FUNCTION_BLOCK EQ_Template (* TEMPLATE for your equipment block, EQ_<Equipment>: copy it under that name, then change what says YOUR OWN, and this comment; keep the rest as it is. An equipment block: the only block that touches this equipment's pins. Skills send it what to switch over a local channel; it switches the outputs (off first, then on), reads the inputs every cycle and reports them to the skills and to OPC UA. One skill holds it at a time; on release or when the module aborts it switches everything off. Technical: A piece of equipment to make your own: one input, one output, one command besides Stop; equipment IO: owns its IO points, writes the output values its holder sends, reads its inputs every cycle and reports changes *)
  (* Standard: 61499-2 *)
  (* Version 0.1, 2026-09-28, Project contributors, AAU Smart Production Lab *)
  PACKAGE stoppering;
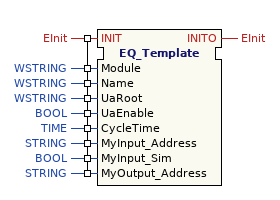
  EVENT_INPUT
    INIT : EInit WITH Module, Name, UaRoot, UaEnable, CycleTime, MyInput_Address, MyInput_Sim, MyOutput_Address; (* Initialise, once at start-up (the INIT chain); takes the values given with it *)
  END_EVENT
  EVENT_OUTPUT
    INITO : EInit; (* Initialised: the next block of the INIT chain goes on *)
  END_EVENT
  VAR_INPUT
    Module : WSTRING; (* The module's name; its local channels are named after it (loc[<Module>/...]) *)
    Name : WSTRING := "Template"; (* YOUR OWN, your equipment's name. The equipment item's name: its local channels and OPC UA folder *)
    UaRoot : WSTRING; (* The module's OPC UA folder, e.g. /Objects/Filling *)
    UaEnable : BOOL; (* Publish on OPC UA *)
    CycleTime : TIME := T#50ms; (* How often the inputs are read *)
    MyInput_Address : STRING; (* YOUR OWN, one per input pin. Where MyInput is: 'gpio[chip:line(:pull_up|:pull_down)(:active_low)]', 'pwm[chip:channel:period_ns]', 'modbus[...]', 'sim', or an IO handle's name; empty: not connected *)
    MyInput_Sim : BOOL := FALSE; (* YOUR OWN, one per input pin. The value of MyInput when simulated (address 'sim') *)
    MyOutput_Address : STRING; (* YOUR OWN, one per output pin. Where MyOutput is: 'gpio[chip:line(:pull_up|:pull_down)(:active_low)]', 'pwm[chip:channel:period_ns]', 'modbus[...]', 'sim', or an IO handle's name; empty: not connected *)
  END_VAR
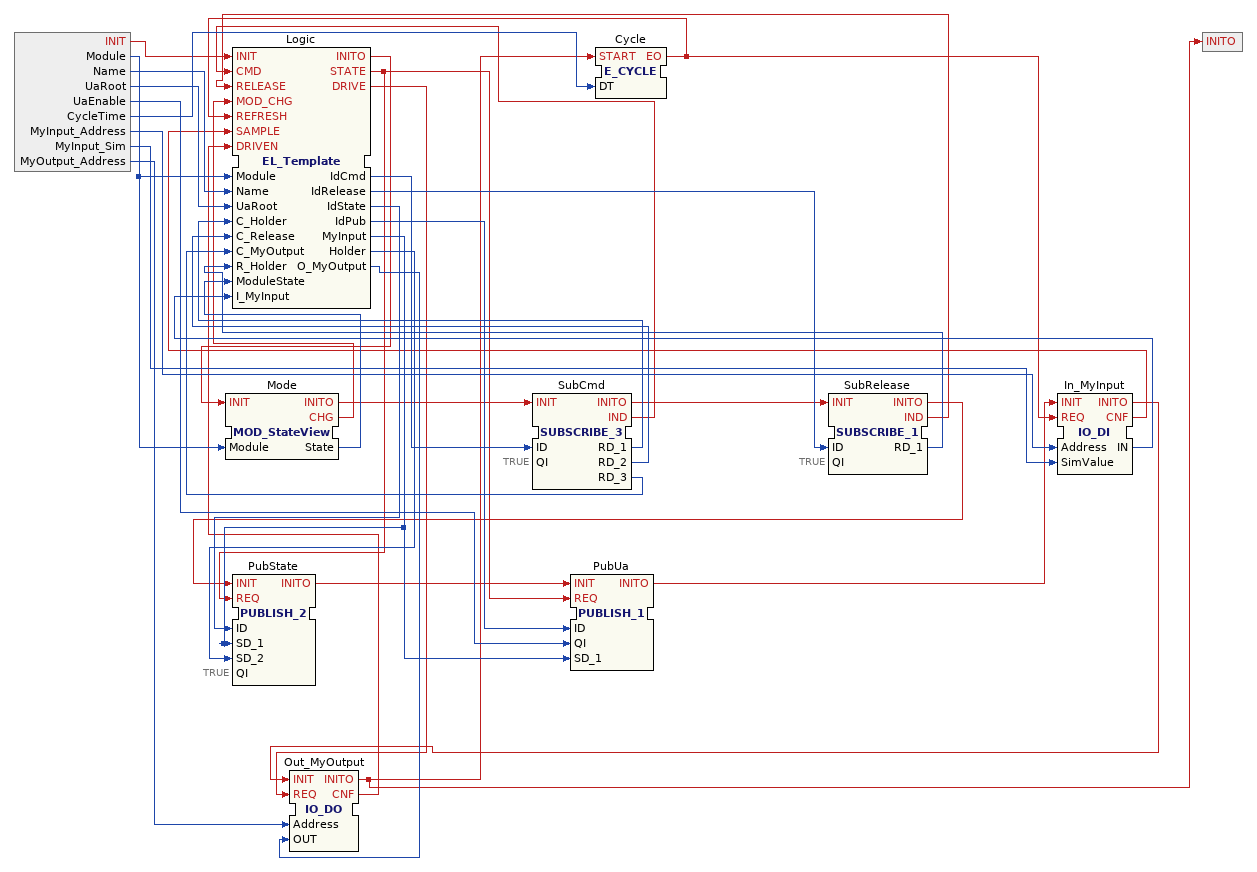
  (* Group Core: One holder at a time, break before make, all off on release or abort; scanned every CycleTime *)
  (* Group Channels: Local channels to and from the skills (cmd, release, state), the module's state, and the inputs over OPC UA *)
  (* Group Inputs: The equipment's sensors: read every cycle, one block per IO point *)
  (* Group Outputs: The equipment's actuators: written on a change and every cycle, one block per IO point *)
  FBS
    Logic : stoppering::EL_Template; (* YOUR OWN, Change Type to your EL_<Equipment>. The equipment's logic (EL_): takes commands from one holder at a time, switches the outputs (off first, then on), switches all off on release or module abort, and reports input changes. *) {SET_ATTRIBUTE(GroupName, Core)}
    Cycle : iec61499::events::E_CYCLE; (* Ticks every cycle so the inputs are read and the outputs refreshed. *) {SET_ATTRIBUTE(GroupName, Core)}
    Mode : modlib::MOD_StateView; (* Watches the module's PackML state, to switch everything off when the module aborts. *) {SET_ATTRIBUTE(GroupName, Channels)}
    SubCmd : iec61499::net::SUBSCRIBE_3(QI := TRUE); (* YOUR OWN, its size: SUBSCRIBE_<outputs + 2>. Receives the commands skills send on this equipment's command channel. *) {SET_ATTRIBUTE(GroupName, Channels)}
    SubRelease : iec61499::net::SUBSCRIBE_1(QI := TRUE); (* Hears the module's release channel: when its holder gives up, everything goes off. *) {SET_ATTRIBUTE(GroupName, Channels)}
    PubState : iec61499::net::PUBLISH_2(QI := TRUE); (* YOUR OWN, its size: PUBLISH_<inputs + 1>. Publishes the inputs and the holder on this equipment's state channel, for the skills. *) {SET_ATTRIBUTE(GroupName, Channels)}
    PubUa : iec61499::net::PUBLISH_1; (* YOUR OWN, its size: PUBLISH_<inputs>; without inputs there is no PubUa. Writes the inputs (and a position, if it keeps one) to OPC UA, below Equipment/<item>. *) {SET_ATTRIBUTE(GroupName, Channels)}
    In_MyInput : modlib::IO_DI; (* YOUR OWN, one per input pin: IO_DI for a switch, IO_AI for an analog input. The pin MyInput: reads the input at MyInput_Address (a Pi pin, Modbus, or simulated). *) {SET_ATTRIBUTE(GroupName, Inputs)}
    Out_MyOutput : modlib::IO_DO; (* YOUR OWN, one per output pin: IO_DO for a switched output, IO_AO for an analog one. The pin MyOutput: switches the output at MyOutput_Address (a Pi pin, Modbus, or simulated). *) {SET_ATTRIBUTE(GroupName, Outputs)}
  END_FBS
  EVENT_CONNECTIONS
    INIT TO Logic.INIT;
    Logic.INITO TO Mode.INIT;
    Mode.INITO TO SubCmd.INIT;
    SubCmd.INITO TO SubRelease.INIT;
    SubRelease.INITO TO PubState.INIT;
    PubState.INITO TO PubUa.INIT;
    PubUa.INITO TO In_MyInput.INIT;
    In_MyInput.INITO TO Out_MyOutput.INIT;
    Out_MyOutput.INITO TO Cycle.START;
    Out_MyOutput.INITO TO INITO;
    SubCmd.IND TO Logic.CMD;
    SubRelease.IND TO Logic.RELEASE;
    Mode.CHG TO Logic.MOD_CHG;
    Cycle.EO TO Logic.REFRESH;
    Cycle.EO TO In_MyInput.REQ;
    In_MyInput.CNF TO Logic.SAMPLE;
    Logic.STATE TO PubState.REQ;
    Logic.STATE TO PubUa.REQ;
    Logic.DRIVE TO Out_MyOutput.REQ;
    Out_MyOutput.CNF TO Logic.DRIVEN;
  END_CONNECTIONS
  DATA_CONNECTIONS
    Module TO Logic.Module;
    Name TO Logic.Name;
    UaRoot TO Logic.UaRoot;
    Module TO Mode.Module;
    Logic.IdCmd TO SubCmd.ID;
    Logic.IdRelease TO SubRelease.ID;
    Logic.IdState TO PubState.ID;
    Logic.IdPub TO PubUa.ID;
    UaEnable TO PubUa.QI;
    CycleTime TO Cycle.DT;
    SubCmd.RD_1 TO Logic.C_Holder;
    SubCmd.RD_2 TO Logic.C_Release;
    SubCmd.RD_3 TO Logic.C_MyOutput;
    SubRelease.RD_1 TO Logic.R_Holder;
    Mode.State TO Logic.ModuleState;
    MyInput_Address TO In_MyInput.Address;
    MyInput_Sim TO In_MyInput.SimValue;
    In_MyInput.IN TO Logic.I_MyInput;
    Logic.MyInput TO PubState.SD_1;
    Logic.MyInput TO PubUa.SD_1;
    Logic.Holder TO PubState.SD_2;
    MyOutput_Address TO Out_MyOutput.Address;
    Logic.O_MyOutput TO Out_MyOutput.OUT;
  END_CONNECTIONS
END_FUNCTION_BLOCK
